(* ================================================================= *)
(*  ST_HandshakeCh                                                   *)
(*  通讯握手通道数据区 - 单通道完整读写区(写+读+诊断)                 *)
(*  版本: V2.0.0  日期: 2026-05-30                                    *)
(*  来源: SysLib/types/                                              *)
(*  变更: 扁平产品数据字段 -> WriteProduct/ReadProduct 嵌入           *)
(* ================================================================= *)

TYPE ST_HandshakeCh :
STRUCT
    Write        : ST_HandshakeBits;   // 写区: 本机->对方 16个Bool信号
    WriteProduct : ST_ProductData;     // 写区产品数据: 本机->对方

    Read         : ST_HandshakeBits;   // 读区: 对方->本机 16个Bool信号
    ReadProduct  : ST_ProductData;     // 读区产品数据: 对方->本机

    CommFault    : BOOL := FALSE;      // 通讯故障综合
    HbTimeout    : BOOL := FALSE;      // 心跳超时
END_STRUCT
END_TYPE
